TEXTLIST TextList_E_Tank_Target
  0 = 'None'
  1 = 'Close'
  2 = 'Open'
  3 = 'Drain'
  4 = 'CIP'
   = ''
END_TEXTLIST

(* stored: Version 1.1.0.1, ProductVersion 3.1.4024.12
   TextList TextList_E_Tank_Target: Id {7337c257-7bcc-4980-8731-40af84e58aad} *)
